SUBAPPLICATION Uebung_159_AX (* Übung zu FsServer: eigener File Server im logiBUS (Gerät B) *)
  (* Standard: 61499-2; Description: Copyright (c) 2026 Meisterschulen am Ostbahnhof This program and the accompanying materials are made available under the terms of the Eclipse Public License 2.0 which is available at https://www.eclipse.org/legal/epl-2.0/ SPDX-License-Identifier: EPL-2.0 *)
  (* Version 1.0, 2026-11-26, Franz Höpfinger, Meisterschulen am Ostbahnhof, initial API and implementation and/or initial documentation *)
  PACKAGE Uebungen;
  IMPORT logiBUS::io::DQ::logiBUS_DO::Output_Q1;
  IMPORT logiBUS::io::DQ::logiBUS_DO::Output_Q2;
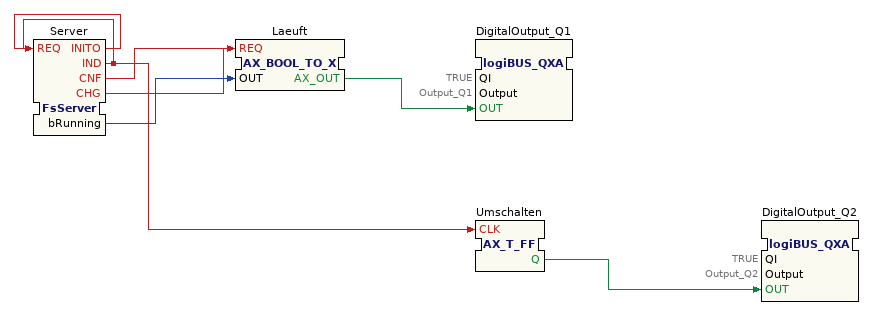
  (* Eigener File Server im logiBUS (FsServer), Gerät B. Gegenstück: Übung 159b auf Gerät A. Einschalten: PART_13_FS = 1 in /data/functionalities.ini, dann Neustart. Optional PART_13_FS_QUOTA_KB (1024) und PART_13_FS_BUS_SHARE (50). Volume \\LOGIBUS\ = /data/fs. Server-CF: NAME-Funktion 61, Herstellercode 1116, Adresse 0xF9. Q1 an = Server läuft (bRunning). Q2 schaltet bei jeder Datei um, die ein Client geschrieben hat (IND). Der Server läuft in der Firmware, auch ohne diesen Baustein. CHG kommt von selbst, wenn sich bRunning, u8Clients oder u8OpenFiles ändert. REQ liest den Status einmal nach INITO und nach jedem IND (u32UsedKB). Watch: bei IND sPath (z. B. /data/fs/IMPORT/test.txt) und u16Lost; nach CNF/CHG u8Clients (1, solange A arbeitet), u8OpenFiles, u32UsedKB, u32QuotaKB. Voraussetzungen: Firmware mit File Server, neue isobus_fs-ELF. Nur ein FsServer pro Gerät. *)
  FBS
    Server : isobus::fs_server::FsServer; (* Volume \\LOGIBUS\ = /data/fs *)
    Laeuft : adapter::conversion::unidirectional::AX_BOOL_TO_X; (* bRunning als AX *)
    DigitalOutput_Q1 : logiBUS::io::DQ::logiBUS_QXA(QI := TRUE, Output := Output_Q1); (* an = Server läuft *)
    Umschalten : adapter::events::unidirectional::AX_T_FF; (* jede geschriebene Datei schaltet Q2 um *)
    DigitalOutput_Q2 : logiBUS::io::DQ::logiBUS_QXA(QI := TRUE, Output := Output_Q2);
  END_FBS
  EVENT_CONNECTIONS
    Server.INITO TO Server.REQ;
    Server.IND TO Server.REQ;
    Server.CNF TO Laeuft.REQ;
    Server.CHG TO Laeuft.REQ;
    Server.IND TO Umschalten.CLK;
  END_CONNECTIONS
  DATA_CONNECTIONS
    Server.bRunning TO Laeuft.OUT;
  END_CONNECTIONS
  ADAPTER_CONNECTIONS
    Laeuft.AX_OUT TO DigitalOutput_Q1.OUT;
    Umschalten.Q TO DigitalOutput_Q2.OUT;
  END_CONNECTIONS
END_SUBAPPLICATION
